(* IEC 61131-3 sources: s22-soft-shell/st_interpret/tests/test_inputs/st_failure/parse_fail, 1 file *)

(* ---- 01_unknown_type.st ---- *)
PROGRAM 01_unknown_type // should error at unknown type
    VAR
	a : Foo;
    END_VAR
	a := 3.1415;
END_PROGRAM
